// TIA Portal V21 export
DATA_BLOCK "IDB_AnaForCounter"   // DB12
// stored: InstanceOfName FB_AnaForCounter, InstanceOfType FB
"FB_AnaForCounter"
   // VAR_INPUT
   //    Limit : Int;
   // END_VAR
   // VAR_OUTPUT
   //    Total : Int;
   // END_VAR
   // VAR
   //    Index : Int;
   // END_VAR
BEGIN
END_DATA_BLOCK
